TYPE ST_RoadRef :
STRUCT
	nMoverCounter: UINT;
	fLength: LREAL;
	pFirstAixs: POINTER TO ST_Axis := null;
	pLastAixs: POINTER TO ST_Axis := null;
	aNode: ARRAY[1..GVL_MC.MAX_MOVER] OF ST_Node;
END_STRUCT
END_TYPE

(* stored: Version 1.1.0.1, ProductVersion 3.1.4024.12
   DUT ST_RoadRef: Id {efe2a556-d5c1-4929-b705-fbd9b88689f3} *)
